Fanuc KAREL source: KT00475.KL

PROGRAM KT00475
%NOLOCKGROUP
VAR
  P1: POSITION
  P2: POSITION
  OUT: XYZWPR
BEGIN
  OUT = P1 : P2
END KT00475
